Fanuc KAREL source: ks00054.KL

-- PROVISIONAL review KL for V1013-1; original PC SHA256 cb9aec1b96bdbe8c5ec60885fbd8f2912ad065d704747e727234f38d202b61ab
-- Incomplete behavior may be omitted. Consult companion uncertainty JSON. Do not deploy.
PROGRAM KS00054
%NOLOCKGROUP
BEGIN
  -- UNRESOLVED_PC offsets 5-13; opcodes 3F,75
  -- UNRESOLVED_PC offsets 18-27; opcodes 3F,75
  -- UNRESOLVED_PC offsets 32-45; opcodes 22,1D,23
  -- UNRESOLVED_PC offsets 50-54; opcodes 7F
END KS00054
